Yaskawa INFORM job: 1KT.JBI

/JOB
//NAME 1KT
//POS
///NPOS 6,6,6,0,0,0
///TOOL 0
///POSTYPE PULSE
///PULSE
C00000=-289,-101140,-84196,3590,-80193,-1939
C00001=-289,-101140,-84196,3590,-80193,-1939
C00002=-103675,52884,19941,-42327,-65457,39225
C00003=-103675,64756,3591,-48976,-53898,45246
C00004=-99503,24499,-40669,-53618,-47781,47266
C00005=-99503,10017,-29148,-45244,-57498,41020
BC00000=570126
BC00001=190240
BC00002=190240
BC00003=190240
BC00004=190240
BC00005=190240
EC00000=-2,-1
EC00001=-2,-1
EC00002=-2,-1
EC00003=-2,-1
EC00004=-2,-1
EC00005=-2,-1
//INST
///DATE 2021/05/18 07:40
///ATTR SC,RW
///GROUP1 RB1,BS1
///GROUP2 ST4
NOP
MOVJ C00000 BC00000 VJ=0.78 PL=0  +MOVJ EC00000 VJ=0.78
MOVJ C00001 BC00001 VJ=0.78 PL=0  +MOVJ EC00001 VJ=0.78
MOVJ C00002 BC00002 VJ=100.00 PL=0  +MOVJ EC00002 VJ=0.78
MOVJ C00003 BC00003 VJ=100.00 PL=0  +MOVJ EC00003 VJ=0.78
ARCON
WVON WEV#(15)
MOVL C00004 BC00004 V=3.3 PL=0  +MOVJ EC00004 VJ=0.78
WVOF
ARCOF
MOVJ C00005 BC00005 VJ=0.78 PL=0  +MOVJ EC00005 VJ=0.78
END
